FUNCTION_BLOCK "LGF_RampCI"
{ S7_Optimized_Access := 'TRUE' }
AUTHOR : Siemens_Digital_Industries
FAMILY : LGF
NAME : LGF_RampCI
   VAR_INPUT
      defaultOutValue : LReal := 0.0;
      contStepNbr : Int := 0;
      contStepTime : Time := T#0MS;
      enDefaulftOutValue : Bool := FALSE;
      start : Bool := FALSE;
      hold : Bool := FALSE;
      continue : Bool := FALSE;
      cyclicOP : Bool := FALSE;
      updateTime : Bool := FALSE;
      reset : Bool := FALSE;
      callOB : OB_CYCLIC;
   END_VAR

   VAR_OUTPUT
      outputValue { ExternalWritable := 'False'} : LReal;
      actTimeTable { ExternalWritable := 'False'} : Bool;
      stepNumber { ExternalWritable := 'False'} : Int;
      remainTime { ExternalWritable := 'False'} : Time;
      totalTime { ExternalWritable := 'False'} : Time;
      remainTotalTime { ExternalWritable := 'False'} : Time;
      error { ExternalWritable := 'False'} : Bool;
      status { ExternalWritable := 'False'} : Word;
      subfunctionStatus { ExternalWritable := 'False'} : Word;
   END_VAR

   VAR_IN_OUT
      setpoints : Array[*] of "LGF_typeRampTimeTable";
   END_VAR

   VAR
      statEndValue { ExternalAccessible := 'False'; ExternalVisible := 'False'; ExternalWritable := 'False'} : LReal;
      statOldValue { ExternalAccessible := 'False'; ExternalVisible := 'False'; ExternalWritable := 'False'} : LReal := 0.0;
      statActualStep { ExternalAccessible := 'False'; ExternalVisible := 'False'; ExternalWritable := 'False'} : Int;
      statActualRestTime { ExternalAccessible := 'False'; ExternalVisible := 'False'; ExternalWritable := 'False'} : Time;
      statTotalTime { ExternalAccessible := 'False'; ExternalVisible := 'False'; ExternalWritable := 'False'} : Time;
      statRestTotalTime { ExternalAccessible := 'False'; ExternalVisible := 'False'; ExternalWritable := 'False'} : Time;
      statStart { ExternalAccessible := 'False'; ExternalVisible := 'False'; ExternalWritable := 'False'} : Bool;
      statTimeTableActiv { ExternalAccessible := 'False'; ExternalVisible := 'False'; ExternalWritable := 'False'} : Bool;
      statStartMem { ExternalAccessible := 'False'; ExternalVisible := 'False'; ExternalWritable := 'False'} : Bool;
      statUpdateTime { ExternalAccessible := 'False'; ExternalVisible := 'False'; ExternalWritable := 'False'} : Bool;
      statReset { ExternalAccessible := 'False'; ExternalVisible := 'False'; ExternalWritable := 'False'} : Bool;
      statResetMem { ExternalAccessible := 'False'; ExternalVisible := 'False'; ExternalWritable := 'False'} : Bool;
   END_VAR

   VAR_TEMP
      tempNewValue : LReal;
      tempIndex : Int;
      tempArrayLowLim : Int;
      tempArrayUpLim : Int;
      tempSampleTime : Time;
      tempCycleTime : UDInt;
      tempCyclePhase : UDInt;
      tempCycleStatus : Word;
      tempReadTimeStatus : Int;
      tempStatus : Word;
   END_VAR

   VAR CONSTANT
      ZERO : Int := 0;
      NO_ERROR : Int := 0;
      RESET_TIME : Time := T#0MS;
      CYCLIC_OB_NOT_AVAILABLE : Word := 16#0000;
      DIMENSION_ONE : UDInt := 1;
      SECOND_IN_MS : UDInt := 1000;
      SUB_STATUS_NO_ERROR : Word := 16#0000;
      STATUS_FINISHED_NO_ERROR : Word := 16#0000;
      STATUS_NO_CALL : Word := 16#7000;
      STATUS_FIRST_CALL : Word := 16#7001;
      STATUS_FURTHER_CALLS : Word := 16#7002;
      ERR_OB_UNAVAILABLE : Word := 16#8200;
      ERR_ARRAY_LOWER_BOUND : Word := 16#8201;
      ERR_QRY_CINT : Word := 16#8400;
   END_VAR


BEGIN
	REGION Block info header
	  //===============================================================================
	  // SIEMENS AG / (c)Copyright 2017
	  //-------------------------------------------------------------------------------
	  // Title:            LGF_RampCI
	  // Comment/Function: Generates a speed curve based on an interpolation point table.
	  // Library/Family:   LGF(Library General Functions)
	  // Author:           Siemens Digital Industry Support
	  // Tested with:      S7-PLCSIM Advanced V2.0 SP1
	  // Engineering:      TIA Portal V15 Update 2
	  // Restrictions:     ENO disabled - error handling done by error and status
	  // Requirements:     PLC (S7-1200 / S7-1500)
	  //-------------------------------------------------------------------------------
	  //=============================================================================
	END_REGION Block info header

	REGION DESCRIPTION
	  (/**/)
	END_REGION DESCRIPTION

	REGION Cycle time
	  // get sample time, according to the cyclic interrupt OB number
	  #tempReadTimeStatus := QRY_CINT(OB_NR := #callOB, CYCLE => #tempCycleTime, PHASE => #tempCyclePhase, STATUS => #tempCycleStatus);
	  #tempCycleTime := #tempCycleTime / #SECOND_IN_MS; // microsecond --> milisecond
	  #tempSampleTime := UDINT_TO_TIME(#tempCycleTime); // Format: TIME

	  #tempStatus := #STATUS_NO_CALL;

	  // Generate error message of the QRY_CINT function
	  IF (#tempReadTimeStatus <> #NO_ERROR) THEN
	    #error := TRUE;
	    #subfunctionStatus := INT_TO_WORD(#tempReadTimeStatus);
	    #status := #ERR_QRY_CINT;
	    RETURN;
	  END_IF;

	  // Generate error message when OB unavailable
	  IF #tempCycleStatus = #CYCLIC_OB_NOT_AVAILABLE THEN
	    #error := TRUE;
	    #status := #ERR_OB_UNAVAILABLE;
	    #subfunctionStatus := #SUB_STATUS_NO_ERROR;
	    RETURN;
	  END_IF;
	END_REGION Cycle time

	REGION Array lower/upper bound
	  #tempArrayLowLim := DINT_TO_INT(LOWER_BOUND(ARR := #setpoints, DIM := #DIMENSION_ONE));
	  #tempArrayUpLim := DINT_TO_INT(UPPER_BOUND(ARR := #setpoints, DIM := #DIMENSION_ONE));

	  IF #tempArrayLowLim <> #ZERO THEN
	    #error := TRUE;
	    #status := #ERR_ARRAY_LOWER_BOUND;
	    #subfunctionStatus := #SUB_STATUS_NO_ERROR;
	    RETURN;
	  END_IF;
	END_REGION Array lower/upper bound

	REGION Function
	  REGION First Call
	    // START by positive edge
	    IF #start AND NOT #statStartMem THEN
	      #tempStatus := #STATUS_FIRST_CALL;
	      #statStart := TRUE;
	      #statTotalTime := #RESET_TIME; // reset total time

	      FOR #tempIndex := #tempArrayLowLim TO #tempArrayUpLim DO // calculate total time
	        #statTotalTime := #statTotalTime + #setpoints[#tempIndex]."time"; // total time
	      END_FOR;
	      #statRestTotalTime := #statTotalTime;
	      #statReset := FALSE;
	    ELSIF NOT #start THEN
	      #error := false;
	      #subfunctionStatus := #SUB_STATUS_NO_ERROR;
	      #status := #STATUS_FINISHED_NO_ERROR;
	    END_IF;
	    // store old value for edge detection
	    #statStartMem := #start;
	  END_REGION First Call

	  REGION Reset
	    // RESET by positiv edge on reset
	    IF #reset AND NOT #statResetMem THEN
	      #tempStatus := #STATUS_FINISHED_NO_ERROR;
	      #statTotalTime := #RESET_TIME; // reset total time

	      FOR #tempIndex := #tempArrayLowLim TO #tempArrayUpLim DO // calculate total time
	        #statTotalTime := #statTotalTime + #setpoints[#tempIndex]."time"; // total time
	      END_FOR;

	      #tempNewValue := #ZERO;                   // output outValue = 0
	      #statRestTotalTime := #statTotalTime;     // update remaining total time
	      #statEndValue := #ZERO;                   // reset statEndValue
	      #statActualStep := #ZERO;                 // reset statActualStep
	      #statActualRestTime := #RESET_TIME;       // reset statActualTime
	      #statStart := TRUE;                       // set start condition
	      #statTimeTableActiv := FALSE;             // reset statTimeTableActive
	      #statReset := TRUE;
	    END_IF;
	    // store old value for edge detection
	    #statResetMem := #reset;
	  END_REGION Reset

	  REGION Operation
	    IF #start AND NOT #statReset THEN
	      // start function ramp soak
	      IF #statStart THEN
	        // Set up start conditions
	        #tempNewValue := #setpoints[#tempArrayLowLim].outputValue;
	        #statEndValue := #setpoints[#tempArrayLowLim + 1].outputValue;
	        #statActualRestTime := #setpoints[#tempArrayLowLim]."time";
	        #statRestTotalTime := #statTotalTime;
	        #statActualStep := 1;
	        #statStart := FALSE;
	        #statTimeTableActiv := TRUE;
	      ELSE
	        IF #hold THEN
	          // Freeze operation
	          #statTimeTableActiv := FALSE;
	          #tempNewValue := #statOldValue;

	          IF #continue THEN
	            // Set up continue conditions
	            // Continue step and remaining time untill continue step
	            #statEndValue := #setpoints[#contStepNbr].outputValue;
	            #statRestTotalTime := #contStepTime;
	            #statActualRestTime := #contStepTime;
	            #statActualStep := #contStepNbr;

	            FOR #tempIndex := #statActualStep TO #tempArrayUpLim DO // calculating remaining total time
	              #statRestTotalTime := #statRestTotalTime + #setpoints[#tempIndex]."time"; // Remaining total time
	            END_FOR;
	          END_IF;
	        ELSE
	          // normal operation
	          // remaining time until actual step
	          IF #statActualRestTime > #tempSampleTime THEN
	            // calculate new output value, if remaining time has not yet expired
	            #tempNewValue := #statOldValue + (#statEndValue - #statOldValue) / DINT_TO_REAL(TIME_TO_DINT(#statActualRestTime)) * UDINT_TO_REAL(#tempCycleTime);
	            // update remaining time till actual step
	            #statActualRestTime := #statActualRestTime - #tempSampleTime;
	            // update remaining total time
	            #statRestTotalTime := #statRestTotalTime - #tempSampleTime;
	          ELSE
	            // remaining actual rest time expired
	            #statActualRestTime := #RESET_TIME;
	            // End of step numbers not reached yet
	            IF #statActualStep < #tempArrayUpLim THEN
	              // set new end value
	              #statEndValue := #setpoints[#statActualStep + 1].outputValue;
	              // set new output value
	              #tempNewValue := #setpoints[#statActualStep].outputValue;
	              // new remaining actual time
	              #statActualRestTime := #setpoints[#statActualStep]."time";
	              #statActualStep := #statActualStep + 1;
	              #statTimeTableActiv := TRUE;
	              #statRestTotalTime := #statRestTotalTime - #tempSampleTime;
	            ELSE
	              // end of step numbers reached
	              #tempStatus := #SUB_STATUS_NO_ERROR;
	              #statRestTotalTime := #RESET_TIME;
	              // cyclic operation
	              IF #cyclicOP THEN
	                #statStart := TRUE;
	                #tempStatus := #STATUS_FURTHER_CALLS;
	              ELSE
	                #statTimeTableActiv := FALSE;
	              END_IF;
	              // set new output value
	              #tempNewValue := #setpoints[#statActualStep].outputValue;
	            END_IF;
	          END_IF;
	        END_IF;
	      END_IF;
	    ELSE
	      #tempNewValue := #ZERO;
	      // time table not active
	      #statTimeTableActiv := FALSE;
	    END_IF;
	  END_REGION Operation

	  REGION Update time
	    // Update total time and remaining total time
	    // Positive edge detection of update time input
	    IF #updateTime AND NOT #statUpdateTime THEN
	      #statTotalTime := #RESET_TIME; // reset total time
	      #statRestTotalTime := #statActualRestTime; // copy remaining actual time to remaining total time

	      FOR #tempIndex := #tempArrayLowLim TO #tempArrayUpLim DO // calculate totel time
	        #statTotalTime := #statTotalTime + #setpoints[#tempIndex]."time"; // total time
	      END_FOR;

	      FOR #tempIndex := #statActualStep TO #tempArrayUpLim DO // calculate remaining total time
	        #statRestTotalTime := #statRestTotalTime + #setpoints[#tempIndex]."time"; // remaining total time
	      END_FOR;
	    END_IF;
	    // store old value for edge detection
	    #statUpdateTime := #updateTime;
	  END_REGION Update time

	  REGION Default output
	    // default value activated: overwrite output by default value
	    IF #enDefaulftOutValue THEN
	      #tempNewValue := #defaultOutValue; // preset output
	      #statTimeTableActiv := FALSE; // timetable not active
	    END_IF;
	  END_REGION Default output
	END_REGION Function

	REGION Write outputs
	  #outputValue := #tempNewValue; // output
	  #statOldValue := #tempNewValue; // store prvious value
	  #actTimeTable := #statTimeTableActiv; //time table active
	  #stepNumber := #statActualStep; // number of acting step
	  #remainTime := #statActualRestTime; // remaining time till actual step
	  #totalTime := #statTotalTime; // total time
	  #remainTotalTime := #statRestTotalTime; //remaining total time

	  #error := #tempStatus.%X15;
	  #status := #tempStatus;
	  #subfunctionStatus := #SUB_STATUS_NO_ERROR;

	  // ENO mechanism is not used
	  ENO := TRUE;
	END_REGION Write outputs

END_FUNCTION_BLOCK